(* IEC 61131-3 sources: plc-st-coding-agent/progress/evidence/full_r8_20261110b/native_evidence/codex_minimax-m27/public-hard-04/1, 1 file *)

(* ---- candidate.st ---- *)
FUNCTION_BLOCK FB
VAR_INPUT
    enqueue  : BOOL;
    dequeue  : BOOL;
    reset    : BOOL;
    capacity : DINT;
END_VAR
VAR_OUTPUT
    elementCount : DINT := 0;
    status       : WORD := 16#0000;
END_VAR
VAR_IN_OUT
    item   : DINT;
    buffer : ARRAY[1..4] OF DINT;
END_VAR
VAR
    head           : DINT := 1;
    tail           : DINT := 1;
    enqueue_prev   : BOOL := FALSE;
    dequeue_prev   : BOOL := FALSE;
END_VAR

// Reset takes priority
IF reset THEN
    elementCount := 0;
    head := 1;
    tail := 1;
    status := 16#0000;
ELSE
    // Idle: no enqueue edge AND no dequeue edge
    IF (enqueue_prev OR NOT enqueue) AND (dequeue_prev OR NOT dequeue) THEN
        status := 16#0000;
    ELSE
        // Rising edge on enqueue
        IF NOT enqueue_prev AND enqueue THEN
            IF elementCount < capacity THEN
                buffer[((tail - 1) MOD capacity) + 1] := item;
                tail := (tail MOD capacity) + 1;
                elementCount := elementCount + 1;
                status := 16#0000;
            ELSE
                status := 16#8002;
            END_IF
        END_IF

        // Rising edge on dequeue
        IF NOT dequeue_prev AND dequeue THEN
            IF elementCount > 0 THEN
                item := buffer[((head - 1) MOD capacity) + 1];
                head := (head MOD capacity) + 1;
                elementCount := elementCount - 1;
                status := 16#0000;
            ELSE
                status := 16#8001;
            END_IF
        END_IF
    END_IF
END_IF

// Update edge detection history at end of scan
enqueue_prev := enqueue;
dequeue_prev := dequeue;
END_FUNCTION_BLOCK
